Universal Robots URScript: step5c_speedj_dryrun_v1.script

# Step5c speedj dry-run quarantine.
# VERSION: 2026-06-13T0041HKT_STEP5C_SPEEDJ_DRYRUN_V1
# GENERATED_AT_LOCAL: 2026-06-13T00:41:36+08:00
# FLOW_TABLE: STEP5_FLOW.md
# STEP5_STAGE_ID: step5c_speedj_dryrun_v1
# STEP5_TABLE_SOURCE: config/step5_stage_table.json
# QUARANTINE_REASON: 2026-06-13 live dry-run moved in the wrong XY/Z direction; DLS/Jacobian mapping is not trusted.
# TP_ROLE: stop_only_quarantine; no motion command, no contact search, no bridge command consumption.
# SAFETY: no speedj, no speedl, no force_mode, no zero_ftsensor(), no TCP/payload write.

def codex_step5c_speedj_dryrun_v1():
  textmsg("codex step5c dry-run quarantine 2026-06-13T0041HKT_STEP5C_SPEEDJ_DRYRUN_V1: DLS/Jacobian mapping wrong; refusing motion")
  write_output_float_register(30, 92.0)
  write_output_float_register(31, 0.0)
  write_output_float_register(35, 29.0)
end

codex_step5c_speedj_dryrun_v1()
